// TIA Portal V19 export
TYPE "ST_USER_BITS_RECIEVE"
   STRUCT
      BUSY : Bool;
      DONE : Bool;
      ERROR : Bool;
      Bit_3 : Bool;
      Bit_4 : Bool;
      Bit_5 : Bool;
      Bit_6 : Bool;
      Bit_7 : Bool;
      Bit_8 : Bool;
      Bit_9 : Bool;
      Bit_10 : Bool;
      Bit_11 : Bool;
      Bit_12 : Bool;
      Bit_13 : Bool;
      Bit_14 : Bool;
      Bit_15 : Bool;
   END_STRUCT;
END_TYPE
